(* IEC 61131-3 sources: PLC_Defuser/Datasets/Water_tank/malicious/mexit, 1 file *)

(* ---- mexit.st ---- *)
FUNCTION_BLOCK valves_handler
  VAR_INPUT
    IN1 : INT;
    IN_TLB1 : INT;
    IN_TLB2 : INT;
  END_VAR
  VAR_OUTPUT
    OUT_MV1 : BOOL;
    OUT_MV2 : BOOL;
  END_VAR
  VAR
    i : INT;
    real_value : INT;
  END_VAR

  real_value :=  IN1 - 5;

  IF real_value <= IN_TLB2 then
    OUT_MV2 := FALSE;
    OUT_MV1 := TRUE;
  end_IF;

  IF real_value >= IN_TLB1 THEN
    OUT_MV2 := TRUE;
    OUT_MV1 := FALSE;
  end_IF;

  i:=0;
  while i<15 do
       OUT_MV2 := FALSE;
       OUT_MV1 := TRUE;
       EXIT;
  end_while;

END_FUNCTION_BLOCK

FUNCTION_BLOCK stop_cycle
  VAR_OUTPUT
    OUT_MV1 : BOOL;
    OUT_MV2 : BOOL;
  END_VAR

  OUT_MV1 := FALSE;
  OUT_MV2 := FALSE;
END_FUNCTION_BLOCK

FUNCTION_BLOCK start_valves
  VAR
    i : INT;
  END_VAR
  VAR_OUTPUT
    OUT_MV2 : BOOL;
    OUT_MV1 : BOOL;
  END_VAR

  i:=0;
  while i<15 do
       OUT_MV2 := TRUE;
       OUT_MV1 := TRUE;

  end_while;
END_FUNCTION_BLOCK

PROGRAM program0
  VAR_INPUT
    TLB2 : INT;
    TLB1 : INT;
    START : BOOL;
    STOP : BOOL;
    VALUE : INT;
  END_VAR
  VAR_OUTPUT
    MV1 : BOOL;
    MV2 : BOOL;
    CYCLE_ON : BOOL;
  END_VAR
  VAR
    valves_handler0 : valves_handler;
    stop_cycle0 : stop_cycle;
    start_valves0 : start_valves;
    _TMP_EQ30_ENO : BOOL;
    _TMP_EQ30_OUT : BOOL;
  END_VAR

  CYCLE_ON := NOT(STOP) AND (CYCLE_ON OR START);
  valves_handler0(EN := CYCLE_ON, IN1 := VALUE, IN_TLB1 := TLB1, IN_TLB2 := TLB2);
  IF valves_handler0.ENO THEN
      MV1 := valves_handler0.OUT_MV1;
  END_IF;
  IF valves_handler0.ENO THEN
      MV2 := valves_handler0.OUT_MV2;
  END_IF;
  stop_cycle0(EN := NOT(CYCLE_ON));
  IF stop_cycle0.ENO THEN
      MV1 := stop_cycle0.OUT_MV1;
  END_IF;
  IF stop_cycle0.ENO THEN
      MV2 := stop_cycle0.OUT_MV2;
  END_IF;
  _TMP_EQ30_OUT := EQ(EN := TRUE, IN1 := VALUE, IN2 := 50, ENO => _TMP_EQ30_ENO);
  start_valves0(EN := _TMP_EQ30_OUT);
  IF start_valves0.ENO THEN
      MV1 := start_valves0.OUT_MV2;
  END_IF;
  IF start_valves0.ENO THEN
      MV2 := start_valves0.OUT_MV1;
  END_IF;
END_PROGRAM

CONFIGURATION Config0

  RESOURCE Res0 ON PLC
    TASK task0(INTERVAL := T#20ms,PRIORITY := 0);
    PROGRAM instance0 WITH task0 : program0;
  END_RESOURCE
END_CONFIGURATION
